FUNCTION_BLOCK FB_SetProductionParams
VAR_INPUT
END_VAR
VAR_OUTPUT
	rCompActualWeight	: REAL;
	iCoun: INT;
	i:INT;
END_VAR
VAR_IN_OUT
	stProdParams		: ST_ProdParams;
	stTriBlender		: ST_TriBlender;
	bTankInProduction	: BOOL;
END_VAR
VAR_INPUT
	iActualWaterAmount	: UINT;
END_VAR


rCompActualWeight:=(TO_REAL(iActualWaterAmount)/100)*stProdParams.arrComponents[i].rCompWeightFor100L;

ACTION act_SetProdVal:

END_ACTION

END_FUNCTION_BLOCK

(* stored: Version 1.1.0.1, ProductVersion 3.1.4024.12
   POU FB_SetProductionParams: Id {ff5743fe-ea81-4a32-8911-c3e1bb7e3f67}, SpecialFunc None
   Action act_SetProdVal: Id {8ebefc7d-d02a-4fa4-a699-82a4ac452993} *)
